FUNCTION "naut_STR_ULINT" : String
{ S7_Optimized_Access := 'TRUE' }
VERSION : 0.1
   VAR_INPUT
      A : ULINT;
   END_VAR
   VAR_TEMP
      s : String;
   END_VAR

BEGIN
	#s := ULINT_TO_STRING(#A);
	IF LEFT(IN := #s, L := 1) = '+' THEN
		#s := DELETE(IN := #s, L := 1, P := 1);
	END_IF;
	#naut_STR_ULINT := #s;
END_FUNCTION
